// TIA Portal V21 export
ORGANIZATION_BLOCK "CallAndCompare"   // OB1, LAD
   VAR_TEMP   // added for the SCL form of the ladder/FBD networks
      _w1 : Bool;
   END_VAR
BEGIN

REGION Network 1: Pump on high level
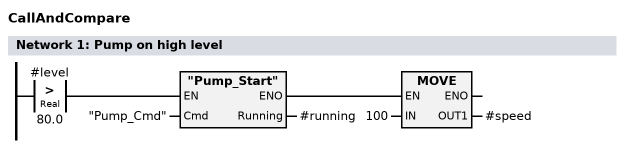
   RUNG wire#powerrail
      { S7_Templates := "SrcType := Real" } GT_Contact(in1 := #level, in2 := 80.0)
      "Pump_Start"(Cmd := "Pump_Cmd", Running => #running)
      Move(in := 100, out1 => #speed)
   END_RUNG
   // the same network as SCL:
   "Pump_Start"(EN := #level > 80.0, Cmd := "Pump_Cmd", Running => #running, ENO => #_w1);
   IF #_w1 THEN #speed := 100; END_IF;
END_REGION
END_ORGANIZATION_BLOCK
